Staubli VAL3: plc.dtx

bool bLifebit = true
bool bReset
bool bSetGun
bool bTosave
public dio dInExcutePainting = {link=3971923C-046E-4FB8-8CDF-8298982DD00B}
dio dInPLCError = {link=0D6C59A5-572E-4845-9D24-D0618D782DD4}
dio dInPowerON = {link=801699AD-0D4E-40AF-A7AF-E7C40311637E}
dio dInResetError = {link=F299EF97-EDDD-4BB8-AA07-719E60051D06}
dio dInStartCycle = {link=842E3CE8-5982-430F-AA8E-B2F701DC178B}
dio dOutCycle = {link=289A5E8D-11F3-4BEB-8FA4-200735E3A2B7}
dio dOutError = {link=79705501-C546-4790-A460-3F340ADFDE5C}
dio dOutEstop = {link=75D4F3C1-C356-4EDA-B423-02C90835EA7D}
dio dOutGunON = {link=734EBAF3-2CA8-4D3F-A8BB-E168C1322725}
dio dOutIsHome = {link=93BF17B5-5C7E-43C6-9C42-3B6025772815}
dio dOutIsPowerd = {link=364EC08F-C077-495B-A954-158507D3C26C}
dio dOutWorkingMode = {link=813E3F4B-A1DE-4C5D-8EAB-0242B6D8A546}
mdesc mNomSpeed
num _bHeavyAlarm
num _nClock = 62473.00582004
num _nNum
num nJointForce[6]
num nLastLib
